// TIA Portal V21 export
DATA_BLOCK "Main_DB"   // DB8
{ S7_Optimized_Access := 'TRUE' }
// stored: MemoryReserve 100
   VAR
      Delay_Time : Time := T#2000ms;
      Delay_done : Bool;
      Delay_in : Bool;
   END_VAR
BEGIN
END_DATA_BLOCK
